(* IEC 61131-3 sources: plc-workbench/outputs/tia_32x4_20261108_results/tasks/01_CUSTOM_01/self_A/details/submissions/3/evaluation/formal, 1 file *)

(* ---- normalized.st ---- *)
FUNCTION_BLOCK FB_ElevatorTarget

   VAR_INPUT
      Enable : BOOL;
      CurrentFloor : INT;
      Direction : INT;
      FullLoad : BOOL;
      CabReq : ARRAY[1 .. 6] OF BOOL;
      HallReq : ARRAY[1 .. 6] OF BOOL;
   END_VAR
   VAR_OUTPUT
      HasTarget : BOOL;
      TargetFloor : INT;
      NextDirection : INT;
   END_VAR
   VAR
      i : INT;
      eligible : BOOL;
      anyEligible : BOOL;
      found : BOOL;
      bestFloor : INT;
      upFloor : INT;
      downFloor : INT;
      absDiff : INT;
      bestAbs : INT;
   END_VAR
VAR_INPUT
WBTEMP_0 : INT;
WBTEMP_1 : BOOL;
WBTEMP_2 : BOOL;
WBTEMP_3 : BOOL;
WBTEMP_4 : INT;
WBTEMP_5 : INT;
WBTEMP_6 : INT;
WBTEMP_7 : INT;
WBTEMP_8 : INT;
END_VAR

i := WBTEMP_0;
eligible := WBTEMP_1;
anyEligible := WBTEMP_2;
found := WBTEMP_3;
bestFloor := WBTEMP_4;
upFloor := WBTEMP_5;
downFloor := WBTEMP_6;
absDiff := WBTEMP_7;
bestAbs := WBTEMP_8;
   HasTarget := FALSE;
   TargetFloor := CurrentFloor;
   NextDirection := 0;

   anyEligible := FALSE;
   FOR i := 1 TO 6 DO
      eligible := CabReq[i] OR (HallReq[i] AND NOT FullLoad);
      IF eligible THEN
         anyEligible := TRUE;
      END_IF;
   END_FOR;

   IF NOT Enable OR NOT anyEligible THEN
      HasTarget := FALSE;
      TargetFloor := CurrentFloor;
      NextDirection := 0;
      RETURN;
   END_IF;

   eligible := CabReq[CurrentFloor] OR (HallReq[CurrentFloor] AND NOT FullLoad);
   IF eligible THEN
      HasTarget := TRUE;
      TargetFloor := CurrentFloor;
      NextDirection := 0;
      RETURN;
   END_IF;

   upFloor := 0;
   downFloor := 0;
   FOR i := 1 TO 6 DO
      eligible := CabReq[i] OR (HallReq[i] AND NOT FullLoad);
      IF eligible AND (i > CurrentFloor) THEN
         IF (upFloor = 0) OR (i < upFloor) THEN
            upFloor := i;
         END_IF;
      END_IF;
      IF eligible AND (i < CurrentFloor) THEN
         IF (downFloor = 0) OR (i > downFloor) THEN
            downFloor := i;
         END_IF;
      END_IF;
   END_FOR;

   bestFloor := CurrentFloor;
   found := FALSE;

   IF Direction = 1 THEN
      IF upFloor > 0 THEN
         bestFloor := upFloor;
         found := TRUE;
      ELSIF downFloor > 0 THEN
         bestFloor := downFloor;
         found := TRUE;
      END_IF;
   ELSIF Direction = -1 THEN
      IF downFloor > 0 THEN
         bestFloor := downFloor;
         found := TRUE;
      ELSIF upFloor > 0 THEN
         bestFloor := upFloor;
         found := TRUE;
      END_IF;
   ELSE
      IF (upFloor > 0) AND (downFloor > 0) THEN
         absDiff := upFloor - CurrentFloor;
         bestAbs := CurrentFloor - downFloor;
         IF absDiff < bestAbs THEN
            bestFloor := upFloor;
            found := TRUE;
         ELSE
            bestFloor := downFloor;
            found := TRUE;
         END_IF;
      ELSIF upFloor > 0 THEN
         bestFloor := upFloor;
         found := TRUE;
      ELSIF downFloor > 0 THEN
         bestFloor := downFloor;
         found := TRUE;
      END_IF;
   END_IF;

   IF found THEN
      HasTarget := TRUE;
      TargetFloor := bestFloor;
      IF bestFloor > CurrentFloor THEN
         NextDirection := 1;
      ELSIF bestFloor < CurrentFloor THEN
         NextDirection := -1;
      ELSE
         NextDirection := 0;
      END_IF;
   ELSE
      HasTarget := FALSE;
      TargetFloor := CurrentFloor;
      NextDirection := 0;
   END_IF;
END_FUNCTION_BLOCK
